Fanuc KAREL source: ko00085.KL

-- PROVISIONAL review KL for V770-1; original PC SHA256 48cea5c80f214abd651b98693ec236a6527235ce887df13b10de6acb47346f20
-- Incomplete behavior may be omitted. Consult companion uncertainty JSON. Do not deploy.
PROGRAM KO00085
%NOLOCKGROUP
BEGIN
  -- UNRESOLVED_PC offsets 5-12; opcodes 9D,23
  -- UNRESOLVED_PC offsets 17-69; opcodes 27,27,49,7E,AD,27,49,7E,AD,22,31,7E,4A
  -- UNRESOLVED_PC offsets 74-78; opcodes 7F
END KO00085
